// TIA Portal V21 export
DATA_BLOCK "LineDb"   // DB43
// stored: AssignedProDiagFB PlantDiag, InstanceOfName Line, InstanceOfType FB
"Line"
BEGIN
END_DATA_BLOCK
